(*
	Immutable snapshot of the identity of one span, created through ContextFactory.buildContext.
	The identifiers are copies, so a context stays valid after the span it came from has ended.
*)
{attribute 'enable_dynamic_creation'}
FUNCTION_BLOCK FB_SpanContext
VAR
	_traceId: FB_TraceId;
	_spanId: FB_SpanId;
	_traceState: POINTER TO FB_TraceState;
	_traceFlags: UDINT;
END_VAR

METHOD _isZero : BOOL
VAR_INPUT
	pBytes: POINTER TO BYTE;
	size: UDINT;
END_VAR
VAR
	i: UDINT;
END_VAR
// bounded by the width of an identifier, at most 16 bytes
_isZero := TRUE;
WHILE i < size DO
	IF pBytes[i] <> 0 THEN
		_isZero := FALSE;
		RETURN;
	END_IF
	i := i + 1;
END_WHILE
END_METHOD

(*
	Releases this context and clears the caller's pointer to it: call it as p^.delete(pSelf:=p).
	pSelf is cleared before the context is freed, so the caller never keeps a dangling pointer.
	A pointer to any other object is refused and left untouched, and nothing is released.
*)
METHOD delete : BOOL
VAR_IN_OUT
	pSelf: POINTER TO FB_SpanContext;
END_VAR
VAR
	_pThis: POINTER TO FB_SpanContext;
END_VAR
_pThis := THIS;
IF pSelf <> _pThis THEN
	RETURN;
END_IF

pSelf := 0;
__DELETE(_pThis);
delete := TRUE;
END_METHOD

//FB_Exit must be implemented explicitly. If there is an implementation, then the
//method is called before the controller removes the code of the function block instance
//(implicit call). The return value is not evaluated.
METHOD FB_Exit: BOOL
VAR_INPUT
    bInCopyCode: BOOL;  // TRUE: the exit method is called in order to leave the instance which will be copied afterwards (online change).
END_VAR
// during an online change the copy keeps the trace state pointer, so it must not be released here
IF NOT bInCopyCode THEN
	THIS^.free();
END_IF
END_METHOD

//FB_Init is always available implicitly and it is used primarily for initialization.
//The return value is not evaluated. For a specific influence, you can also declare the
//methods explicitly and provide additional code there with the standard initialization
//code. You can evaluate the return value.
METHOD FB_Init: BOOL
VAR_INPUT
    bInitRetains: BOOL; // TRUE: the retain variables are initialized (reset warm / reset cold)
    bInCopyCode: BOOL;  // TRUE: the instance will be copied to the copy code afterward (online change)
	pTraceId: POINTER TO FB_TraceId;  // copied
	pSpanId: POINTER TO FB_SpanId;  // copied
	pTraceState: POINTER TO FB_TraceState;  // ownership transfers to the context; 0 means none
	traceFlags: UDINT;
END_VAR
(*
Allocation and argument checks are done by ContextFactory and not the context itself,
that way a new context never gets allocated if building it fails.
The identity is not validated; producers are responsible for what they build.
*)
IF pTraceId <> 0 THEN
	MEMCPY(ADR(THIS^._traceId.bytes), ADR(pTraceId^.bytes), SIZEOF(THIS^._traceId.bytes));
END_IF
IF pSpanId <> 0 THEN
	MEMCPY(ADR(THIS^._spanId.bytes), ADR(pSpanId^.bytes), SIZEOF(THIS^._spanId.bytes));
END_IF
THIS^._traceState := pTraceState;
THIS^._traceFlags := traceFlags;
FB_Init := TRUE;
END_METHOD

//FB_Reinit is called after the instance has been copied during an online change.
//The return value is not evaluated.
METHOD FB_Reinit: BOOL
// nothing to fix up: the trace state lives on the heap and does not move with the instance,
// and no member points back into this instance
FB_Reinit := TRUE;
END_METHOD

(*
	Releases the trace state and clears the identity. Safe to call more than once.
*)
METHOD free
IF THIS^._traceState <> 0 THEN
	THIS^._traceState^.delete(pSelf:=THIS^._traceState);
END_IF
THIS^._traceId.free();
THIS^._spanId.free();
THIS^._traceFlags := 0;
END_METHOD

(*
	TRUE only when remoteness is known and the span is remote, meaning the context was
	extracted from a carrier rather than produced by a local tracer.
	FALSE covers both "known local" and "not known".
*)
METHOD isRemote : BOOL
isRemote := (THIS^._traceFlags AND TO_UDINT(E_SpanFlags.SPAN_FLAGS_CONTEXT_HAS_IS_REMOTE_MASK)) <> 0
	AND (THIS^._traceFlags AND TO_UDINT(E_SpanFlags.SPAN_FLAGS_CONTEXT_IS_REMOTE_MASK)) <> 0;
END_METHOD

(*
	TRUE if and only if both the trace ID and the span ID are non-zero.
*)
METHOD isValid : BOOL
isValid := NOT THIS^._isZero(pBytes := ADR(THIS^._traceId.bytes), size := SIZEOF(THIS^._traceId.bytes))
	AND NOT THIS^._isZero(pBytes := ADR(THIS^._spanId.bytes), size := SIZEOF(THIS^._spanId.bytes));
END_METHOD

PROPERTY spanId : REFERENCE TO FB_SpanId
GET
spanId REF= THIS^._spanId;
END_GET
END_PROPERTY

PROPERTY traceFlags : UDINT
GET
traceFlags := THIS^._traceFlags;
END_GET
END_PROPERTY

PROPERTY traceId : REFERENCE TO FB_TraceId
GET
traceId REF= THIS^._traceId;
END_GET
END_PROPERTY

// borrowed; 0 when the context carries no trace state. The context owns and releases it.
PROPERTY traceState : POINTER TO FB_TraceState
GET
traceState := THIS^._traceState;
END_GET
END_PROPERTY

END_FUNCTION_BLOCK

(* stored: Version 1.1.0.1
   POU FB_SpanContext: Id {cb3780ad-42f4-466e-beb9-8fb650ce5375}, SpecialFunc None
   Method _isZero: Id {ba7fa559-df6e-42aa-a334-d206d09748cb}
   Method delete: Id {091fc591-8b0e-413b-bd89-1ac90e00a59c}
   Method FB_Exit: Id {bd5ef56d-2d7a-4740-8b81-5bb55127c6a7}
   Method FB_Init: Id {9cd3ddcd-9701-47d5-891f-b3d3b0d18b1c}
   Method FB_Reinit: Id {27b958f9-35d6-4d2e-b40f-bc7f83136759}
   Method free: Id {12adc99d-389b-4fc1-8440-eecf17b8fe3b}
   Method isRemote: Id {c2cb054f-a30e-4b73-affe-ebe12a7607ce}
   Method isValid: Id {467f115c-472e-426d-89cb-b2ff80cda960}
   Property spanId: Id {a28cd319-5be4-48bd-881a-0d2ddbc180b1}
   Get Get: Id {1bfe45b3-fd8c-4c30-8c82-2291a189b428}
   Property traceFlags: Id {2bc93955-48b9-47fb-b0b8-96e6e5f5550a}
   Get Get: Id {ee7720d6-e477-45e8-9c31-d91a133f6889}
   Property traceId: Id {656b1a0e-13e9-4281-a9d1-ceb9792387a5}
   Get Get: Id {02d984f9-7cf1-42ca-854c-98c4361f860d}
   Property traceState: Id {c41eee4f-4355-47a1-8e2c-83ab681255ff}
   Get Get: Id {2bdadfbd-495f-4b25-b861-a6f5573bba15} *)
